{attribute 'pack_mode' := '1'}
TYPE ST_ScheduleDaily_V1 :
STRUCT
	Name : STRING(20);
	Priority : UDINT;
	StartDate : UDINT;
	EndDate : UDINT;
	Works : ARRAY[0..9] OF ST_ScheduleWork_V1;
END_STRUCT
END_TYPE

(* stored: Version 1.1.0.1, ProductVersion 3.1.4024.15
   DUT ST_ScheduleDaily_V1: Id {c90a2b4a-b601-4a30-a9a8-76350db2573d} *)
